// TIA Portal V18 export
TYPE "Process_Gap"
   STRUCT
      ProcessGapActive : Bool;
      ModezoneGap { S7_SetPoint := 'True'} : Array[1.."ModeZone_Setup_Const"] of "Modezone_Gap";
   END_STRUCT;
END_TYPE
